Universal Robots PolyScope program: EdgeProg.urp

Program EdgeProg (createdIn=3.0.0 lastSavedIn=3.0.0 directory=/programs installation=default)
Robot Program (runOnlyOnce=true motionType=MoveJ speed=1.047198 acceleration=1.396263 useActiveTCP=false)
  'Program generated by RoboDK v6.0.7 for ABB IRB 120-3/0.6 on XX/XX/XXXX 18:00:00'
  'Using nominal kinematics.'
  'Using Ref. Frame Edge: p[0.100500, -0.200250, 0.300125, 0.547381, -0.295318, 0.260260]'
  'Using TCP Tool Edge: p[-0.001500, 0.002250, 0.099875, -1.759988, 1.759988, 0.729011]'
  Script: set_tcp(p[-0.001500, 0.002250, 0.099875, -1.759988, 1.759988, 0.729011])
  Script: movej([-0.087266, -0.087266, 0.261799, 0.174533, 0.698132, -0.174533],1.20000,0.58177,0,0.0000)
  MoveJ speed 33.35 deg/s, acceleration 68.75 deg/s^2 (useActiveTCP=true)
    Waypoint Waypoint_1: TCP in base x=-265.419 y=-512.444 z=406.972 mm, rx=0.0789 ry=2.1217 rz=0.5281 rad; joints [-5, -5, 15, 10, 40, -10] deg; flange x=-251.297 y=-472.118 z=316.657 mm, rx=0.4756 ry=0.1811 rz=-1.4344 rad
  MoveL speed 123 mm/s, acceleration 1200 mm/s^2 (useActiveTCP=true)
    Waypoint Waypoint_2: motionParameters(blendRadius=0.013); TCP in base x=-752.411 y=-79.146 z=724.974 mm, rx=0.208 ry=1.5218 rz=-0.4854 rad; joints [-5, -5, 15, 10, 40, -10] deg; flange x=-692.318 y=-122.405 z=657.894 mm, rx=0.3644 ry=-0.9259 rz=-1.8089 rad
  Halt
  Wait Sleep waitTime=1.234
  Popup Message (haltProgram=false message=A long message with "quotes", 'apostrophes' & symbols: <>[]{}()=+-*/%;#@! and more text to make it longer than eighty characters)
  'Comment with ; semicolon'
  Set DigitalOutput pin=Gripper; digitalValue=ON
  Set DigitalOutput pin=digital_out[12]; digitalValue=0
  Set DigitalOutput pin=Pressure; digitalValue=1
  Wait DigitalInput pin=PartPresent; digitalValue=1
  Wait DigitalInput pin=digital_in[get_standard_digital_in(7)]; digitalValue=1
  Call DoSomething
  Script: x = 1
  Script: movej([0.349066, -0.174533, 0.349066, 0.000000, 0.523599, 0.000000],1.20000,0.58177,0,0.0000)
SubProgram  [hidden by the author, left out]
SubProgram DoSomething [hidden by the author, left out]
